            num nDelay = 1
            num nMoveType = 1
            num nPercentage
            num nSigValue
        pointRx pPointRx[2] = {x=379.796411, y=595.987022, z=1351.538711, rx=1.401068, ry=1.345217, rz=-178.109847, shoulder=lefty, elbow=epositive, wrist=wpositive}
        string sID
      [9]
        bool bMarked
        jointRx jJointRx = {j1=39.880437, j2=-6.575361, j3=82.0777309, j4=-177.996823, j5=75.37833, j6=-38.47744}
        pointRx pInter
        paraItem pParaItem
          [0]
            bool bSafePoint
            ifItem iIfItem
              [0]
                bool bANDOR[2]
                num nSigIndex[3]
                num nSigType[3]
                num nValue[3]
            mdesc mMdesc = {leave=0}
            num nActionIndex = 41
            num nDelay = 1
            num nMoveType = 1
            num nPercentage
            num nSigValue
        pointRx pPointRx[2] = {x=379.796362, y=520.320173, z=1238.0913856, rx=1.402674, ry=1.344381, rz=-178.109837, shoulder=lefty, elbow=epositive, wrist=wpositive}
        string sID
      [10]
        bool bMarked
        jointRx jJointRx = {j1=41.803306, j2=-6.517095, j3=92.330616, j4=-178.0541377, j5=85.747638, j6=-40.0393449}
        pointRx pInter
        paraItem pParaItem
          [0]
            bool bSafePoint
            ifItem iIfItem
              [0]
                bool bANDOR[2]
                num nSigIndex[3]
                num nSigType[3]
                num nValue[3]
            mdesc mMdesc = {leave=0}
            num nActionIndex = 41
            num nDelay = 1
            num nMoveType = 1
            num nPercentage
            num nSigValue
        pointRx pPointRx[2] = {x=379.334807, y=543.604553, z=1140.610387, rx=1.401253, ry=1.344273, rz=-178.109295, shoulder=lefty, elbow=epositive, wrist=wpositive}
        string sID
      [11]
        bool bMarked
        jointRx jJointRx = {j1=41.782649, j2=-6.517552, j3=100.0447353, j4=-178.0556323, j5=93.456121, j6=-39.757291}
        pointRx pInter
        paraItem pParaItem
          [0]
            bool bSafePoint
            ifItem iIfItem
              [0]
                bool bANDOR[2]
                num nSigIndex[3]
                num nSigType[3]
                num nValue[3]
            mdesc mMdesc = {leave=0}
            num nActionIndex = 41
            num nDelay = 1
            num nMoveType = 1
            num nPercentage
            num nSigValue
        pointRx pPointRx[2] = {x=379.796355, y=543.749536, z=1066.621752, rx=1.401483, ry=1.344544, rz=-178.109518, shoulder=lefty, elbow=epositive, wrist=wpositive}
        string sID
      [12]
        bool bMarked
        jointRx jJointRx = {j1=34.795273, j2=-10.731385, j3=113.971463, j4=-178.0324342, j5=102.926788, j6=-32.442855}
        pointRx pInter
        paraItem pParaItem
          [0]
            bool bSafePoint
            ifItem iIfItem
              [0]
                bool bANDOR[2]
                num nSigIndex[3]
                num nSigType[3]
                num nValue[3]
            mdesc mMdesc = {leave=0}
            num nActionIndex = 41
            num nDelay = 1
            num nMoveType = 1
            num nPercentage
            num nSigValue
        pointRx pPointRx[2] = {x=384.534447, y=467.177264, z=968.97583, rx=1.400551, ry=1.345316, rz=-178.109467, shoulder=lefty, elbow=epositive, wrist=wpositive}
        string sID
      [13]
        bool bMarked
        jointRx jJointRx = {j1=21.426698, j2=-20.557567, j3=119.218666, j4=-178.186954, j5=97.91655, j6=-19.25856}
        pointRx pInter
        paraItem pParaItem
          [0]
            bool bSafePoint
            ifItem iIfItem
              [0]
                bool bANDOR[2]
                num nSigIndex[3]
                num nSigType[3]
                num nValue[3]
            mdesc mMdesc = {leave=0}
            num nActionIndex = 41
            num nDelay = 1
            num nMoveType = 1
            num nPercentage
            num nSigValue
        pointRx pPointRx[2] = {x=379.796362, y=344.491625, z=989.0258456, rx=1.401479, ry=1.345115, rz=-178.109716, shoulder=lefty, elbow=epositive, wrist=wpositive}
        string sID
      [14]
        bool bMarked
        jointRx jJointRx = {j1=21.573037, j2=-21.112859, j3=107.354759, j4=-178.196288, j5=85.509411, j6=-19.796082}
        pointRx pInter
        paraItem pParaItem
          [0]
            bool bSafePoint
            ifItem iIfItem
              [0]
                bool bANDOR[2]
                num nSigIndex[3]
                num nSigType[3]
                num nValue[3]
            mdesc mMdesc = {leave=0}
            num nActionIndex = 41
            num nDelay = 1
            num nMoveType = 1
            num nPercentage
            num nSigValue
        pointRx pPointRx[2] = {x=379.796366, y=345.634221, z=1106.178535, rx=1.40246, ry=1.344064, rz=-178.109758, shoulder=lefty, elbow=epositive, wrist=wpositive}
        string sID
      [15]
        bool bMarked
        jointRx jJointRx = {j1=55.916319, j2=-32.435037, j3=81.208272, j4=-180.529582, j5=50.673289, j6=-143.736818}
        pointRx pInter
        paraItem pParaItem
          [0]
            bool bSafePoint
            ifItem iIfItem
              [0]
                bool bANDOR[2]
                num nSigIndex[3]
                num nSigType[3]
                num nValue[3]
            mdesc mMdesc = {leave=0}
            num nActionIndex = 41
            num nDelay = 1
            num nMoveType = 1
            num nPercentage
            num nSigValue
        pointRx pPointRx[2] = {x=213.314986, y=180.947183, z=1388.164351, rx=1.343298, ry=-1.403323, rz=91.85354, shoulder=lefty, elbow=epositive, wrist=wpositive}
        string sID
      [16]
        bool bMarked
        jointRx jJointRx = {j1=51.328619, j2=-33.392172, j3=100.816411, j4=-180.357794, j5=69.338541, j6=-141.673567}
        pointRx pInter
        paraItem pParaItem
          [0]
            bool bSafePoint
            ifItem iIfItem
              [0]
                bool bANDOR[2]
                num nSigIndex[3]
                num nSigType[3]
                num nValue[3]
            mdesc mMdesc = {leave=0}
            num nActionIndex = 41
            num nDelay = 1
            num nMoveType = 1
            num nPercentage
            num nSigValue
        pointRx pPointRx[2] = {x=282.275825, y=237.105347, z=1232.303049, rx=1.285321, ry=-1.457217, rz=89.539558, shoulder=lefty, elbow=epositive, wrist=wpositive}
        string sID
      [17]
        bool bMarked
        jointRx jJointRx = {j1=51.324147, j2=-34.916794, j3=105.550027, j4=-180.350309, j5=72.547076, j6=-141.690388}
        pointRx pInter
        paraItem pParaItem
          [0]
            bool bSafePoint
            ifItem iIfItem
              [0]
                bool bANDOR[2]
                num nSigIndex[3]
                num nSigType[3]
                num nValue[3]
            mdesc mMdesc = {leave=0}
            num nActionIndex = 41
            num nDelay = 1
            num nMoveType = 1
            num nPercentage
            num nSigValue
        pointRx pPointRx[2] = {x=282.310453, y=237.105448, z=1196.0721274, rx=1.285273, ry=-1.456601, rz=89.539451, shoulder=lefty, elbow=epositive, wrist=wpositive}
        string sID
      [18]
        bool bMarked
        jointRx jJointRx = {j1=47.711546, j2=-35.77088, j3=112.0332318, j4=-180.218474, j5=78.193659, j6=-138.139834}
        pointRx pInter
        paraItem pParaItem
          [0]
            bool bSafePoint
            ifItem iIfItem
              [0]
                bool bANDOR[2]
                num nSigIndex[3]
                num nSigType[3]
                num nValue[3]
            mdesc mMdesc = {leave=0}
            num nActionIndex = 41
            num nDelay = 1
            num nMoveType = 1
            num nPercentage
            num nSigValue
        pointRx pPointRx[2] = {x=304.164757, y=234.823085, z=1139.987435, rx=1.285005, ry=-1.457553, rz=89.539753, shoulder=lefty, elbow=epositive, wrist=wpositive}
        string sID
      [19]
        bool bMarked
        jointRx jJointRx = {j1=57.172461, j2=-20.295318, j3=103.584374, j4=-181.910796, j5=82.86872, j6=-234.262378}
        pointRx pInter
        paraItem pParaItem
          [0]
            bool bSafePoint
            ifItem iIfItem
              [0]
                bool bANDOR[2]
                num nSigIndex[3]
                num nSigType[3]
                num nValue[3]
            mdesc mMdesc = {leave=0}
            num nActionIndex = 41
            num nDelay = 1
            num nMoveType = 1
            num nPercentage
            num nSigValue
        pointRx pPointRx[2] = {x=180.349472, y=237.105491, z=1136.925483, rx=-1.3845, ry=-1.363197, rz=2.663332, shoulder=lefty, elbow=epositive, wrist=wpositive}
        string sID
      [20]
        bool bMarked
        jointRx jJointRx = {j1=58.963813, j2=-17.899384, j3=106.645873, j4=-181.882945, j5=88.263458, j6=-236.241021}
        pointRx pInter
        paraItem pParaItem
          [0]
            bool bSafePoint
            ifItem iIfItem
              [0]
                bool bANDOR[2]
                num nSigIndex[3]
                num nSigType[3]
                num nValue[3]
            mdesc mMdesc = {leave=0}
            num nActionIndex = 41
            num nDelay = 1
            num nMoveType = 1
            num nPercentage
            num nSigValue
        pointRx pPointRx[2] = {x=180.349453, y=262.820622, z=1091.52565, rx=-1.38517, ry=-1.363097, rz=2.657182, shoulder=lefty, elbow=epositive, wrist=wpositive}
        string sID
      [21]
        bool bMarked
        jointRx jJointRx = {j1=11.381472, j2=-45.430894, j3=114.894163, j4=-226.110043, j5=69.582957, j6=-170.981239}
        pointRx pInter
        paraItem pParaItem
          [0]
            bool bSafePoint
            ifItem iIfItem
              [0]
                bool bANDOR[2]
                num nSigIndex[3]
                num nSigType[3]
                num nValue[3]
            mdesc mMdesc = {leave=0}
            num nActionIndex = 41
            num nDelay = 1
            num nMoveType = 1
            num nPercentage
            num nSigValue
        pointRx pPointRx[2] = {x=180.349761, y=382.492889, z=1091.525435, rx=-43.00473097, ry=-2.0901953, rz=2.639534, shoulder=lefty, elbow=epositive, wrist=wpositive}
        string sID
      [22]
        bool bMarked
        jointRx jJointRx = {j1=16.208393, j2=-31.573324, j3=103.438513, j4=-221.00332249, j5=83.760859, j6=-158.676963}
        pointRx pInter
        paraItem pParaItem
          [0]
            bool bSafePoint
            ifItem iIfItem
              [0]
                bool bANDOR[2]
                num nSigIndex[3]
                num nSigType[3]
                num nValue[3]
            mdesc mMdesc = {leave=0}
            num nActionIndex = 41
            num nDelay = 1
            num nMoveType = 1
            num nPercentage
            num nSigValue
        pointRx pPointRx[2] = {x=157.842425, y=384.0224699, z=1151.632552, rx=-38.308759, ry=-17.884638, rz=22.19937, shoulder=lefty, elbow=epositive, wrist=wpositive}
        string sID
      [23]
        bool bMarked
        jointRx jJointRx = {j1=18.812847, j2=-31.349268, j3=104.945814, j4=-221.438921, j5=83.42439, j6=-161.706803}
        pointRx pInter
        paraItem pParaItem
          [0]
            bool bSafePoint
            ifItem iIfItem
              [0]
                bool bANDOR[2]
                num nSigIndex[3]
                num nSigType[3]
                num nValue[3]
            mdesc mMdesc = {leave=0}
            num nActionIndex = 41
            num nDelay = 1
            num nMoveType = 1
            num nPercentage
            num nSigValue
        pointRx pPointRx[2] = {x=157.667732, y=398.947608, z=1136.779994, rx=-38.309247, ry=-17.885155, rz=22.199699, shoulder=lefty, elbow=epositive, wrist=wpositive}
        string sID
      [24]
        bool bMarked
        jointRx jJointRx = {j1=96.0913, j2=-31.728358, j3=114.0722837, j4=-202.614442, j5=94.0603229, j6=-157.248945}
        pointRx pInter
        paraItem pParaItem
          [0]
            bool bSafePoint
            ifItem iIfItem
              [0]
                bool bANDOR[2]
                num nSigIndex[3]
                num nSigType[3]
                num nValue[3]
            mdesc mMdesc = {leave=0}
            num nActionIndex = 41
            num nDelay = 1
            num nMoveType = 1
            num nPercentage
            num nSigValue
        pointRx pPointRx[2] = {x=-173.392959, y=252.540582, z=1108.905783, rx=14.434003, ry=-21.15753, rz=120.829292, shoulder=lefty, elbow=epositive, wrist=wpositive}
        string sID
      [25]
        bool bMarked
        jointRx jJointRx = {j1=166.142444, j2=11.119509, j3=74.56791, j4=-164.63285, j5=110.70051, j6=-117.214853}
        pointRx pInter
        paraItem pParaItem
          [0]
            bool bSafePoint
            ifItem iIfItem
              [0]
                bool bANDOR[2]
                num nSigIndex[3]
                num nSigType[3]
                num nValue[3]
            mdesc mMdesc = {leave=0}
            num nActionIndex = 41
            num nDelay = 1
            num nMoveType = 1
            num nPercentage
            num nSigValue
        pointRx pPointRx[2] = {x=-512.796929, y=314.598166, z=1094.722813, rx=-9.112922, ry=27.868894, rz=-131.0635766, shoulder=lefty, elbow=epositive, wrist=wpositive}
        string sID
      [26]
        bool bMarked
        jointRx jJointRx = {j1=13.104952, j2=-46.838042, j3=98.098651, j4=-173.383208, j5=52.299423, j6=-42.459137}
        pointRx pInter
        paraItem pParaItem
          [0]
            bool bSafePoint
            ifItem iIfItem
              [0]
                bool bANDOR[2]
                num nSigIndex[3]
                num nSigType[3]
                num nValue[3]
            mdesc mMdesc = {leave=0}
            num nActionIndex = 41
            num nDelay = 1
            num nMoveType = 1
            num nPercentage
            num nSigValue
        pointRx pPointRx[2] = {x=172.0214078, y=163.423356, z=1296.555569, rx=5.287932, ry=0.356736, rz=154.726012, shoulder=lefty, elbow=epositive, wrist=wpositive}
        string sID
      [27]
        bool bMarked
        jointRx jJointRx = {j1=-0.746077, j2=38.654193, j3=103.0610419, j4=-179.633028, j5=123.454226, j6=8.386419}
        pointRx pInter
        paraItem pParaItem
          [0]
            bool bSafePoint
            ifItem iIfItem
              [0]
                bool bANDOR[2]
                num nSigIndex[3]
                num nSigType[3]
                num nValue[3]
            mdesc mMdesc = {leave=10}
            num nActionIndex = 41
            num nDelay = 1
            num nMoveType = 1
            num nPercentage
            num nSigValue
        pointRx pPointRx[2] = {x=872.305806, y=193.820048, z=536.464849, rx=0.56853, ry=18.254398, rz=-172.702509, shoulder=lefty, elbow=epositive, wrist=wpositive}
        string sID
      [28]
        bool bMarked
        jointRx jJointRx = {j1=-0.746077, j2=38.654194, j3=103.0610414, j4=-179.633029, j5=123.454226, j6=8.386419}
        pointRx pInter
        paraItem pParaItem
          [0]
            bool bSafePoint
            ifItem iIfItem
              [0]
                bool bANDOR[2]
                num nSigIndex[3]
                num nSigType[3]
                num nValue[3]
            mdesc mMdesc = {leave=0}
            num nActionIndex = 71
            num nDelay = 1
            num nMoveType = 4
            num nPercentage
            num nSigValue
        pointRx pPointRx[2] = {x=872.305806, y=193.820048, z=536.464849, rx=0.56853, ry=18.254398, rz=-172.702509, shoulder=lefty, elbow=epositive, wrist=wpositive}
        string sID
      [29]
        bool bMarked
        jointRx jJointRx = {j1=-0.746077, j2=38.654194, j3=103.0610414, j4=-179.633029, j5=123.454226, j6=8.386419}
        pointRx pInter
        paraItem pParaItem
          [0]
            bool bSafePoint
            ifItem iIfItem
              [0]
                bool bANDOR[2]
                num nSigIndex[3]
                num nSigType[3]
                num nValue[3]
            mdesc mMdesc = {leave=0}
            num nActionIndex = 70
            num nDelay = 1
            num nMoveType = 4
            num nPercentage
            num nSigValue = 1
        pointRx pPointRx[2] = {x=872.305806, y=193.820048, z=536.464849, rx=0.56853, ry=18.254398, rz=-172.702509, shoulder=lefty, elbow=epositive, wrist=wpositive}
        string sID
      [30]
        bool bMarked
        jointRx jJointRx = {j1=-0.746077, j2=38.654194, j3=103.0610414, j4=-179.633029, j5=123.454226, j6=8.386419}
        pointRx pInter
        paraItem pParaItem
          [0]
            bool bSafePoint
            ifItem iIfItem
              [0]
                bool bANDOR[2]
                num nSigIndex[3]
                num nSigType[3]
                num nValue[3]
            mdesc mMdesc = {leave=0}
            num nActionIndex = 70
            num nDelay = 1
            num nMoveType = 3
            num nPercentage
            num nSigValue = 1
        pointRx pPointRx[2] = {x=872.305806, y=193.820048, z=536.464849, rx=0.56853, ry=18.254398, rz=-172.702509, shoulder=lefty, elbow=epositive, wrist=wpositive}
        string sID
    string sID
  [PR02-WashPATH2]
    num nFrameIndex
    num nMoveID
    num nToolIndex
    pointItem pPointItem[118]
      [0]
        bool bMarked
        jointRx jJointRx = {j1=1.472874, j2=128.415304, j3=-142.718421, j4=-10.676075, j5=-13.610921, j6=92.673149}
        pointRx pInter
        paraItem pParaItem
          [0]
            bool bSafePoint
            ifItem iIfItem
              [0]
                bool bANDOR[2]
                num nSigIndex[3]
                num nSigType[3]
                num nValue[3]
            mdesc mMdesc
            num nActionIndex = 60
            num nDelay = 1
            num nMoveType = 7
            num nPercentage
            num nSigValue = 1
        pointRx pPointRx[2] = {x=91.326194, y=-43.762939, z=599.882275, rx=-88.611323, ry=-173.490167, rz=-62.0834554, shoulder=lefty, elbow=enegative, wrist=wnegative}
        string sID
      [1]
        bool bMarked
        jointRx jJointRx = {j1=-0.746435, j2=38.656305, j3=103.0621354, j4=-179.633633, j5=123.453008, j6=8.386286}
        pointRx pInter
        paraItem pParaItem
          [0]
            bool bSafePoint
            ifItem iIfItem
              [0]
                bool bANDOR[2]
                num nSigIndex[3]
                num nSigType[3]
                num nValue[3]
            mdesc mMdesc = {leave=0}
            num nActionIndex = 60
            num nDelay = 1
            num nMoveType = 1
            num nPercentage
            num nSigValue = 1
        pointRx pPointRx[2] = {x=872.340958, y=193.819324, z=536.420305, rx=0.568193, ry=18.258826, rz=-172.70256, shoulder=lefty, elbow=epositive, wrist=wpositive}
        string sID
      [2]
        bool bMarked
        jointRx jJointRx = {j1=13.421878, j2=-4.818376, j3=127.477265, j4=-178.119237, j5=122.0948701, j6=-9.80116}
        pointRx pInter
        paraItem pParaItem
          [0]
            bool bSafePoint
            ifItem iIfItem
              [0]
                bool bANDOR[2]
                num nSigIndex[3]
                num nSigType[3]
                num nValue[3]
            mdesc mMdesc = {leave=0}
            num nActionIndex = 60
            num nDelay = 1
            num nMoveType = 1
            num nPercentage
            num nSigValue = 1
        pointRx pPointRx[2] = {x=448.783781, y=302.866041, z=805.255089, rx=1.42221, ry=0.904693, rz=-177.39771, shoulder=lefty, elbow=epositive, wrist=wpositive}
        string sID
      [3]
        bool bMarked
        jointRx jJointRx = {j1=-44.645904, j2=7.328511, j3=115.0443755, j4=-179.561776, j5=120.728528, j6=47.488337}
        pointRx pInter
        paraItem pParaItem
          [0]
            bool bSafePoint
            ifItem iIfItem
              [0]
                bool bANDOR[2]
                num nSigIndex[3]
                num nSigType[3]
                num nValue[3]
            mdesc mMdesc = {leave=0}
            num nActionIndex = 60
            num nDelay = 1
            num nMoveType = 1
            num nPercentage
            num nSigValue = 1
        pointRx pPointRx[2] = {x=448.783853, y=-225.927858, z=805.255091, rx=1.423155, ry=0.904518, rz=-177.398128, shoulder=lefty, elbow=epositive, wrist=wpositive}
        string sID
      [4]
        bool bMarked
        jointRx jJointRx = {j1=-60.278459, j2=-4.417844, j3=115.214708, j4=-181.80285, j5=110.802192, j6=150.0409807}
        pointRx pInter
        paraItem pParaItem
          [0]
            bool bSafePoint
            ifItem iIfItem
              [0]
                bool bANDOR[2]
                num nSigIndex[3]
                num nSigType[3]
                num nValue[3]
            mdesc mMdesc = {leave=0}
            num nActionIndex = 60
            num nDelay = 1
            num nMoveType = 1
            num nPercentage
            num nSigValue = 1
        pointRx pPointRx[2] = {x=159.335469, y=-423.920881, z=907.0568085, rx=-0.848529, ry=1.45622, rz=-89.586458, shoulder=lefty, elbow=epositive, wrist=wpositive}
        string sID
      [5]
        bool bMarked
        jointRx jJointRx = {j1=-71.457668, j2=-10.942695, j3=120.893936, j4=-181.757898, j5=110.283853, j6=161.255103}
        pointRx pInter
        paraItem pParaItem
          [0]
            bool bSafePoint
            ifItem iIfItem
              [0]
                bool bANDOR[2]
                num nSigIndex[3]
                num nSigType[3]
                num nValue[3]
            mdesc mMdesc = {leave=0}
            num nActionIndex = 60
            num nDelay = 1
            num nMoveType = 1
            num nPercentage
            num nSigValue = 1
        pointRx pPointRx[2] = {x=52.814992, y=-423.885575, z=907.0568224, rx=-0.848102, ry=1.454685, rz=-89.587129, shoulder=lefty, elbow=epositive, wrist=wpositive}
        string sID
      [6]
        bool bMarked
        jointRx jJointRx = {j1=-84.239451, j2=-15.195174, j3=124.219334, j4=-181.627917, j5=109.714573, j6=174.101598}
        pointRx pInter
        paraItem pParaItem
          [0]
            bool bSafePoint
            ifItem iIfItem
              [0]
                bool bANDOR[2]
                num nSigIndex[3]
                num nSigType[3]
                num nValue[3]
            mdesc mMdesc = {leave=0}
            num nActionIndex = 60
            num nDelay = 1
            num nMoveType = 1
            num nPercentage
            num nSigValue = 1
        pointRx pPointRx[2] = {x=-50.911318, y=-423.885576, z=907.0568257, rx=-0.848073, ry=1.4547, rz=-89.587134, shoulder=lefty, elbow=epositive, wrist=wpositive}
        string sID
      [7]
        bool bMarked
        jointRx jJointRx = {j1=-98.383773, j2=-16.506532, j3=125.186653, j4=-181.397639, j5=109.725834, j6=188.326149}
        pointRx pInter
        paraItem pParaItem
          [0]
            bool bSafePoint
            ifItem iIfItem
              [0]
                bool bANDOR[2]
                num nSigIndex[3]
                num nSigType[3]
                num nValue[3]
            mdesc mMdesc = {leave=0}
            num nActionIndex = 60
            num nDelay = 1
            num nMoveType = 1
            num nPercentage
            num nSigValue = 1
        pointRx pPointRx[2] = {x=-157.789841, y=-423.885562, z=907.0568281, rx=-0.848066, ry=1.4548, rz=-89.587112, shoulder=lefty, elbow=epositive, wrist=wpositive}
        string sID
      [8]
        bool bMarked
        jointRx jJointRx = {j1=-112.0278043, j2=-14.344006, j3=123.577475, j4=-181.102464, j5=110.562296, j6=202.0554572}
        pointRx pInter
        paraItem pParaItem
          [0]
            bool bSafePoint
            ifItem iIfItem
              [0]
                bool bANDOR[2]
                num nSigIndex[3]
                num nSigType[3]
                num nValue[3]
            mdesc mMdesc = {leave=0}
            num nActionIndex = 60
            num nDelay = 1
            num nMoveType = 1
            num nPercentage
            num nSigValue = 1
        pointRx pPointRx[2] = {x=-265.4041, y=-423.885563, z=907.056825, rx=-0.847933, ry=1.456541, rz=-89.586315, shoulder=lefty, elbow=epositive, wrist=wpositive}
        string sID
      [9]
        bool bMarked
        jointRx jJointRx = {j1=-123.571629, j2=-9.344784, j3=119.568416, j4=-180.800027, j5=111.732577, j6=213.687233}
        pointRx pInter
        paraItem pParaItem
          [0]
            bool bSafePoint
            ifItem iIfItem
              [0]
                bool bANDOR[2]
                num nSigIndex[3]
                num nSigType[3]
                num nValue[3]
            mdesc mMdesc = {leave=0}
            num nActionIndex = 60
            num nDelay = 1
            num nMoveType = 1
            num nPercentage
            num nSigValue = 1
        pointRx pPointRx[2] = {x=-371.195573, y=-423.885577, z=907.0568224, rx=-0.847959, ry=1.454646, rz=-89.587183, shoulder=lefty, elbow=epositive, wrist=wpositive}
        string sID
      [10]
        bool bMarked
        jointRx jJointRx = {j1=-132.987781, j2=-2.32091, j3=113.237219, j4=-180.526229, j5=112.527397, j6=223.195107}
        pointRx pInter
        paraItem pParaItem
          [0]
            bool bSafePoint
            ifItem iIfItem
              [0]
                bool bANDOR[2]
                num nSigIndex[3]
                num nSigType[3]
                num nValue[3]
            mdesc mMdesc = {leave=0}
            num nActionIndex = 60
            num nDelay = 1
            num nMoveType = 1
            num nPercentage
            num nSigValue = 1
        pointRx pPointRx[2] = {x=-478.725239, y=-423.885573, z=907.0568161, rx=-0.847819, ry=1.454622, rz=-89.587133, shoulder=lefty, elbow=epositive, wrist=wpositive}
        string sID
      [11]
        bool bMarked
        jointRx jJointRx = {j1=-137.536891, j2=0.364167, j3=110.596819, j4=-180.386169, j5=112.606426, j6=227.795437}
        pointRx pInter
        paraItem pParaItem
          [0]
            bool bSafePoint
            ifItem iIfItem
              [0]
                bool bANDOR[2]
                num nSigIndex[3]
                num nSigType[3]
                num nValue[3]
            mdesc mMdesc = {leave=0}
            num nActionIndex = 60
            num nDelay = 1
            num nMoveType = 1
            num nPercentage
            num nSigValue = 1
        pointRx pPointRx[2] = {x=-529.0764983, y=-411.740053, z=907.0568193, rx=-0.848313, ry=1.454843, rz=-89.587359, shoulder=lefty, elbow=epositive, wrist=wpositive}
        string sID
      [12]
        bool bMarked
        jointRx jJointRx = {j1=-132.35753, j2=-10.0229591, j3=120.136433, j4=-180.542512, j5=111.720654, j6=222.565935}
        pointRx pInter
        paraItem pParaItem
          [0]
            bool bSafePoint
            ifItem iIfItem
              [0]
                bool bANDOR[2]
                num nSigIndex[3]
                num nSigType[3]
                num nValue[3]
            mdesc mMdesc = {leave=0}
            num nActionIndex = 60
            num nDelay = 1
            num nMoveType = 1
            num nPercentage
            num nSigValue = 1
        pointRx pPointRx[2] = {x=-430.774932, y=-380.176303, z=907.0568091, rx=-0.848827, ry=1.455835, rz=-89.587105, shoulder=lefty, elbow=epositive, wrist=wpositive}
        string sID
      [13]
        bool bMarked
        jointRx jJointRx = {j1=-118.807255, j2=-18.339875, j3=126.49453, j4=-180.921153, j5=109.59715, j6=208.9121}
        pointRx pInter
        paraItem pParaItem
          [0]
            bool bSafePoint
            ifItem iIfItem
              [0]
                bool bANDOR[2]
                num nSigIndex[3]
                num nSigType[3]
                num nValue[3]
            mdesc mMdesc = {leave=0}
            num nActionIndex = 60
            num nDelay = 1
            num nMoveType = 1
            num nPercentage
            num nSigValue = 1
        pointRx pPointRx[2] = {x=-300.995578, y=-380.211371, z=907.0568212, rx=-0.847914, ry=1.456586, rz=-89.586337, shoulder=lefty, elbow=epositive, wrist=wpositive}
        string sID
      [14]
        bool bMarked
        jointRx jJointRx = {j1=-101.602024, j2=-22.421109, j3=129.221385, j4=-181.320362, j5=107.919298, j6=191.610896}
        pointRx pInter
        paraItem pParaItem
          [0]
            bool bSafePoint
            ifItem iIfItem
              [0]
                bool bANDOR[2]
                num nSigIndex[3]
                num nSigType[3]
                num nValue[3]
            mdesc mMdesc = {leave=0}
            num nActionIndex = 60
            num nDelay = 1
            num nMoveType = 1
            num nPercentage
            num nSigValue = 1
        pointRx pPointRx[2] = {x=-173.307357, y=-380.211369, z=907.0568274, rx=-0.847854, ry=1.456568, rz=-89.586358, shoulder=lefty, elbow=epositive, wrist=wpositive}
        string sID
      [15]
        bool bMarked
        jointRx jJointRx = {j1=-83.0907973, j2=-20.866813, j3=128.212142, j4=-181.627255, j5=108.00511422, j6=172.999356}
        pointRx pInter
        paraItem pParaItem
          [0]
            bool bSafePoint
            ifItem iIfItem
              [0]
                bool bANDOR[2]
                num nSigIndex[3]
                num nSigType[3]
                num nValue[3]
            mdesc mMdesc = {leave=0}
            num nActionIndex = 60
            num nDelay = 1
            num nMoveType = 1
            num nPercentage
            num nSigValue = 1
        pointRx pPointRx[2] = {x=-47.315982, y=-380.211387, z=907.056824, rx=-0.847929, ry=1.456122, rz=-89.586559, shoulder=lefty, elbow=epositive, wrist=wpositive}
        string sID
      [16]
        bool bMarked
        jointRx jJointRx = {j1=-66.0904757, j2=-14.194712, j3=123.463577, j4=-181.776403, j5=109.444961, j6=155.904397}
        pointRx pInter
        paraItem pParaItem
          [0]
            bool bSafePoint
            ifItem iIfItem
              [0]
                bool bANDOR[2]
                num nSigIndex[3]
                num nSigType[3]
                num nValue[3]
            mdesc mMdesc = {leave=0}
            num nActionIndex = 60
            num nDelay = 1
            num nMoveType = 1
            num nPercentage
            num nSigValue = 1
        pointRx pPointRx[2] = {x=82.0110787, y=-380.211384, z=907.0568184, rx=-0.847913, ry=1.456404, rz=-89.586467, shoulder=lefty, elbow=epositive, wrist=wpositive}
        string sID
      [17]
        bool bMarked
        jointRx jJointRx = {j1=-56.975917, j2=-4.42927, j3=115.225272, j4=-181.798703, j5=110.703168, j6=146.741231}
        pointRx pInter
        paraItem pParaItem
          [0]
            bool bSafePoint
            ifItem iIfItem
              [0]
                bool bANDOR[2]
                num nSigIndex[3]
                num nSigType[3]
                num nValue[3]
            mdesc mMdesc = {leave=0}
            num nActionIndex = 60
            num nDelay = 1
            num nMoveType = 1
            num nPercentage
            num nSigValue = 1
        pointRx pPointRx[2] = {x=183.647044, y=-405.622287, z=907.05681, rx=-0.847156, ry=1.456129, rz=-89.586622, shoulder=lefty, elbow=epositive, wrist=wpositive}
        string sID
      [18]
        bool bMarked
        jointRx jJointRx = {j1=-53.343407, j2=-3.133018, j3=114.0121449, j4=-181.789883, j5=110.680859, j6=143.111047}
        pointRx pInter
        paraItem pParaItem
          [0]
            bool bSafePoint
            ifItem iIfItem
              [0]
                bool bANDOR[2]
                num nSigIndex[3]
                num nSigType[3]
                num nValue[3]
            mdesc mMdesc = {leave=0}
            num nActionIndex = 60
            num nDelay = 1
            num nMoveType = 1
            num nPercentage
            num nSigValue = 1
        pointRx pPointRx[2] = {x=215.747782, y=-392.804263, z=907.0568113, rx=-0.848298, ry=1.456111, rz=-89.586519, shoulder=lefty, elbow=epositive, wrist=wpositive}
        string sID
      [19]
        bool bMarked
        jointRx jJointRx = {j1=-31.769864, j2=-17.771615, j3=126.0947542, j4=-181.560446, j5=107.525433, j6=121.69219}
        pointRx pInter
        paraItem pParaItem
          [0]
            bool bSafePoint
            ifItem iIfItem
              [0]
                bool bANDOR[2]
                num nSigIndex[3]
                num nSigType[3]
                num nValue[3]
            mdesc mMdesc = {leave=0}
            num nActionIndex = 60
            num nDelay = 1
            num nMoveType = 1
            num nPercentage
            num nSigValue = 1
        pointRx pPointRx[2] = {x=238.277852, y=-170.574116, z=907.0568198, rx=-0.848582, ry=1.456262, rz=-89.586608, shoulder=lefty, elbow=epositive, wrist=wpositive}
        string sID
      [20]
        bool bMarked
        jointRx jJointRx = {j1=-33.0616256, j2=-27.634624, j3=132.351778, j4=-181.551134, j5=103.955202, j6=123.0799891}
        pointRx pInter
        paraItem pParaItem
          [0]
            bool bSafePoint
            ifItem iIfItem
              [0]
                bool bANDOR[2]
                num nSigIndex[3]
                num nSigType[3]
                num nValue[3]
            mdesc mMdesc = {leave=0}
            num nActionIndex = 60
            num nDelay = 1
            num nMoveType = 1
            num nPercentage
            num nSigValue = 1
        pointRx pPointRx[2] = {x=175.936032, y=-141.263692, z=907.0568162, rx=-0.848923, ry=1.45551, rz=-89.586745, shoulder=lefty, elbow=epositive, wrist=wpositive}
        string sID
      [21]
        bool bMarked
        jointRx jJointRx = {j1=-46.679029, j2=-38.679088, j3=137.790309, j4=-181.659354, j5=98.725516, j6=136.824211}
        pointRx pInter
        paraItem pParaItem
          [0]
            bool bSafePoint
            ifItem iIfItem
              [0]
                bool bANDOR[2]
                num nSigIndex[3]
                num nSigType[3]
                num nValue[3]
            mdesc mMdesc = {leave=0}
            num nActionIndex = 60
            num nDelay = 1
            num nMoveType = 1
            num nPercentage
            num nSigValue = 1
        pointRx pPointRx[2] = {x=84.172629, y=-162.0462482, z=907.0568202, rx=-0.847558, ry=1.455278, rz=-89.58679, shoulder=lefty, elbow=epositive, wrist=wpositive}
        string sID
      [22]
        bool bMarked
        jointRx jJointRx = {j1=-74.173892, j2=-54.901318, j3=143.26089, j4=-181.630942, j5=88.779079, j6=164.61695}
        pointRx pInter
        paraItem pParaItem
          [0]
            bool bSafePoint
            ifItem iIfItem
              [0]
                bool bANDOR[2]
                num nSigIndex[3]
                num nSigType[3]
                num nValue[3]
            mdesc mMdesc = {leave=0}
            num nActionIndex = 60
            num nDelay = 1
            num nMoveType = 1
            num nPercentage
            num nSigValue = 1
        pointRx pPointRx[2] = {x=-44.604354, y=-162.0461536, z=907.0568118, rx=-0.847894, ry=1.454483, rz=-89.586903, shoulder=lefty, elbow=epositive, wrist=wpositive}
        string sID
      [23]
        bool bMarked
        jointRx jJointRx = {j1=-116.822113, j2=-59.877841, j3=144.419733, j4=-180.917751, j5=85.955845, j6=207.300383}
        pointRx pInter
        paraItem pParaItem
          [0]
            bool bSafePoint
            ifItem iIfItem
              [0]
                bool bANDOR[2]
                num nSigIndex[3]
                num nSigType[3]
                num nValue[3]
            mdesc mMdesc = {leave=0}
            num nActionIndex = 60
            num nDelay = 1
            num nMoveType = 1
            num nPercentage
            num nSigValue = 1
        pointRx pPointRx[2] = {x=-174.555607, y=-162.0463469, z=907.0568299, rx=-0.848322, ry=1.454721, rz=-89.586982, shoulder=lefty, elbow=epositive, wrist=wpositive}
        string sID
      [24]
        bool bMarked
        jointRx jJointRx = {j1=-145.38456, j2=-48.183629, j3=141.324497, j4=-180.128817, j5=94.81986, j6=235.777806}
        pointRx pInter
        paraItem pParaItem
          [0]
            bool bSafePoint
            ifItem iIfItem
              [0]
                bool bANDOR[2]
                num nSigIndex[3]
                num nSigType[3]
                num nValue[3]
            mdesc mMdesc = {leave=0}
            num nActionIndex = 60
            num nDelay = 1
            num nMoveType = 1
            num nPercentage
            num nSigValue = 1
        pointRx pPointRx[2] = {x=-302.7407, y=-162.0462705, z=907.0568236, rx=-0.848311, ry=1.454665, rz=-89.587042, shoulder=lefty, elbow=epositive, wrist=wpositive}
        string sID
      [25]
        bool bMarked
        jointRx jJointRx = {j1=-157.976861, j2=-30.800178, j3=134.0695528, j4=-179.751099, j5=104.935628, j6=248.439783}
        pointRx pInter
        paraItem pParaItem
          [0]
            bool bSafePoint
            ifItem iIfItem
              [0]
                bool bANDOR[2]
                num nSigIndex[3]
                num nSigType[3]
                num nValue[3]
            mdesc mMdesc = {leave=0}
